FUNCTION_BLOCK "FB_StlC_049"
TITLE = STL call WRITE_BIG
{ S7_Optimized_Access := 'TRUE' }
VERSION : 0.1
   VAR_INPUT
      a : Bool;
      i1 : Int;
      i2 : Int;
      di1 : DInt;
      r1 : Real;
      w1 : Word;
      dw1 : DWord;
      b1 : Byte;
      u1 : UInt;
      ud1 : UDInt;
   END_VAR

   VAR_OUTPUT
      q : Bool;
      io : Int;
      dio : DInt;
      ro : Real;
      wo : Word;
      dwo : DWord;
      bo : Byte;
      udo : UDInt;
   END_VAR

   VAR_IN_OUT
      v : Variant;
      arrs : Array[*] of Int;
      pos : DInt;
   END_VAR

   VAR
      src : Array[0..9] of Int;
      dst : Array[0..9] of Int;
      bits : Array[0..31] of Bool;
      bytes : Array[0..9] of Byte;
      err {InstructionName := 'ErrorStruct'; LibVersion := '1.0'} : ErrorStruct;
      rt : LReal;
      tim {InstructionName := 'IEC_TIMER'; LibVersion := '1.0'} : IEC_TIMER;
      words : Array[0..3] of Word;
   END_VAR


BEGIN
NETWORK
TITLE = 049 WRITE_BIG
      CALL WRITE_BIG
      {src_type := 'Int', dst_type := 'Variant'}
      (  src_variable                := #i1 ,
         OUT                         := #io ,
         dest_array                  := #bytes ,
         pos                         := #pos
      );
END_FUNCTION_BLOCK

